Fanuc KAREL source: kd00054.KL

-- PROVISIONAL review KL for V1013-1; original PC SHA256 ace4c5ae55d14bbc955efe60db36277c8d552eb0675a44ef077f401a73eb9d87
-- Incomplete behavior may be omitted. Consult companion uncertainty JSON. Do not deploy.
PROGRAM KD00054
%NOLOCKGROUP
VAR
  I : INTEGER
  J : INTEGER
  B : BOOLEAN
  R : REAL
  S : STRING[80]
BEGIN
  -- UNRESOLVED_PC offsets 5-28; opcodes 9D,81,18,9D,1B,9D,12,22,2E,13,04
  -- UNRESOLVED_PC offsets 33-37; opcodes 7F
END KD00054
